// TIA Portal V18 export
// export: Created 2026-11-25T00:00:00.0000000Z, ExportSetting WithDefaults
Connection "Connection_PLC"  Driver=SIMATIC S7 1500, InterfaceType=Ethernet
  AreaPointer   AreaPointerType=Coordination
  AreaPointer   AreaPointerType=DateTime
  AreaPointer   AreaPointerType=DateTimereturn
  AreaPointer   AreaPointerType=EventId
  AreaPointer   AreaPointerType=FieldbusReadmailbox
  AreaPointer   AreaPointerType=FieldbusWritemailbox
  AreaPointer   AreaPointerType=HmiIdentification
  AreaPointer   AreaPointerType=Jobmailbox
  AreaPointer   AreaPointerType=ProjectId
  AreaPointer   AreaPointerType=ScreenNumber
  AreaPointer   AreaPointerType=TagManagement
